(* PLC project Vn_op_expt, Beckhoff Automation GmbH TwinCAT PLC Control 3.5.13.21 *)
(* stored: creationDateTime 1970-01-01T00:00:00 *)

PROGRAM Vn_op_expt

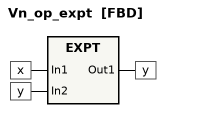
(* FBD diagram, written out as Structured Text *)
y := EXPT(x, y);
END_PROGRAM
